// TwinCAT 3 PLC project MQTT_PLC_TEST
// ProgramVersion: 3.1.4024.0
// libraries:
//   Tc2_Standard, * (Beckhoff Automation GmbH)
//   Tc2_System, * (Beckhoff Automation GmbH)
//   Tc2_Utilities, * (Beckhoff Automation GmbH)
//   Tc3_IotBase, * (Beckhoff Automation GmbH)
//   Tc3_Module, * (Beckhoff Automation GmbH)
// project tree:
//   / GlobalTextList.TcGTLO, PlcTask.TcTTO
//   GVLs/ GVL_Visu.TcGVL, GVL_Mqtt.TcGVL
//   POUs/ MAIN.TcPOU
//   VISUs/ PannenkoekenDashboard.TcVIS
// real-time tasks:
//   TASK PlcTask: cycle T#10ms, priority 20, ADS port 350
// I/O:
//   DEVICE Device 1 (EtherCAT) (disabled), AmsNetId 199.4.42.250.2.1
//     Term 1 (EK1200) [EK1200-5000 EtherCAT Power supply (2A E-Bus)]
//       Term 2 (EL1008) [EL1008 8Ch. Dig. Input 24V, 3ms]
//       Term 3 (EL2008) [EL2008 8Ch. Dig. Output 24V, 0.5A]
//       Term 4 (EL3062) [EL3062 2Ch. Ana. Input 0-10V]
//       Term 5 (EL4002) [EL4002 2Ch. Ana. Output 0-10V, 12bit]
//       Term 6 (EK1110) [EK1110 EtherCAT extension]

CONFIGURATION MQTT_PLC_TEST
    RESOURCE PLC ON TwinCAT3
        TASK PlcTask(INTERVAL := T#10ms, PRIORITY := 20);
        PROGRAM MAIN WITH PlcTask : MAIN;
    END_RESOURCE
END_CONFIGURATION

// ---- GVLs/GVL_Visu.TcGVL
{attribute 'qualified_only'}
VAR_GLOBAL
    // Robot Arm
    sRobotState        : STRING(10);   // idle, moving, error
    nRobotColor        : DWORD;        // kleur voor rectangle/LED
    bRobotCmdSentPulse : BOOL;         // pulse indicator
    bRobotStateParseError : BOOL;      // parse fout indicator
END_VAR

// ---- GVLs/GVL_Mqtt.TcGVL
VAR_GLOBAL CONSTANT
    c_sMqttHost           : STRING(63) := '192.168.0.197';
    c_nMqttPort           : UINT := 1883;

    c_sTopicRobotCmd      : STRING(127) := 'pancake/robot/cmd';
    c_sTopicRobotState    : STRING(127) := 'pancake/robot/state';
    c_sTopicRobotError    : STRING(127) := 'pancake/robot/error';
    c_sTopicConveyorCmd   : STRING(127) := 'pancake/conveyor/cmd';
    c_sTopicConveyorState : STRING(127) := 'pancake/conveyor/state';
    c_sTopicConveyorError : STRING(127) := 'pancake/conveyor/error';
END_VAR

VAR_GLOBAL
    bMqttEnable                : BOOL := TRUE;
    bMqttConnected             : BOOL;
    bMqttError                 : BOOL;
    sMqttStatus                : STRING(127);

    sRobotState                : STRING(31) := 'unknown';
    bRobotStateUpdated         : BOOL;
    bRobotStateParseError      : BOOL;

    sConveyorCmdRx             : STRING(31);
    bConveyorCmdUpdated        : BOOL;
    sConveyorState             : STRING(31) := 'stopped';
    sConveyorStatePublished    : STRING(31);
    bConveyorStateSentPulse    : BOOL;
    sConveyorErrorText         : STRING(127);
    bConveyorErrorSentPulse    : BOOL;
    sConveyorItem              : STRING(31);
    bConveyorItemPresent       : BOOL;
    bConveyorItemUpdated       : BOOL;

    sRobotErrorRx              : STRING(127);
    bRobotErrorUpdated         : BOOL;

    sRobotCmdRequest           : STRING(31);
    bRobotCmdRequestPulse      : BOOL;
    sRobotCmdPending           : STRING(31);
    sRobotCmdSent              : STRING(31);
    bRobotCmdSentPulse         : BOOL;

    sCoordinatorState          : STRING(31);
    sLastRxTopic               : STRING(127);
    sLastRxPayload             : STRING(255);

    bCmdPick                   : BOOL;
    bCmdPlace                  : BOOL;
    bCmdHome                   : BOOL;
    bCmdStop                   : BOOL;
END_VAR

// ---- POUs/MAIN.TcPOU
PROGRAM MAIN
VAR
END_VAR

END_PROGRAM

// ---- GlobalTextList.TcGTLO
TEXTLIST GlobalTextList
  14 = 'Broker Host'
  78 = 'Broker Port'
  184 = 'Connected'
  631 = 'E-STOP'
  815 = 'E-STOPS'
  297 = 'Enable MQTT'
  818 = 'Error'
  717 = 'Mixer'
  369 = 'MQTT Broker'
  28 = 'MQTT Monitor'
  441 = 'Robot Arm'
  964 = 'Robot State'
  282 = 'S'
  632 = 'Status'
  865 = 'Transportband'
END_TEXTLIST

// ---- VISUs/PannenkoekenDashboard.TcVIS
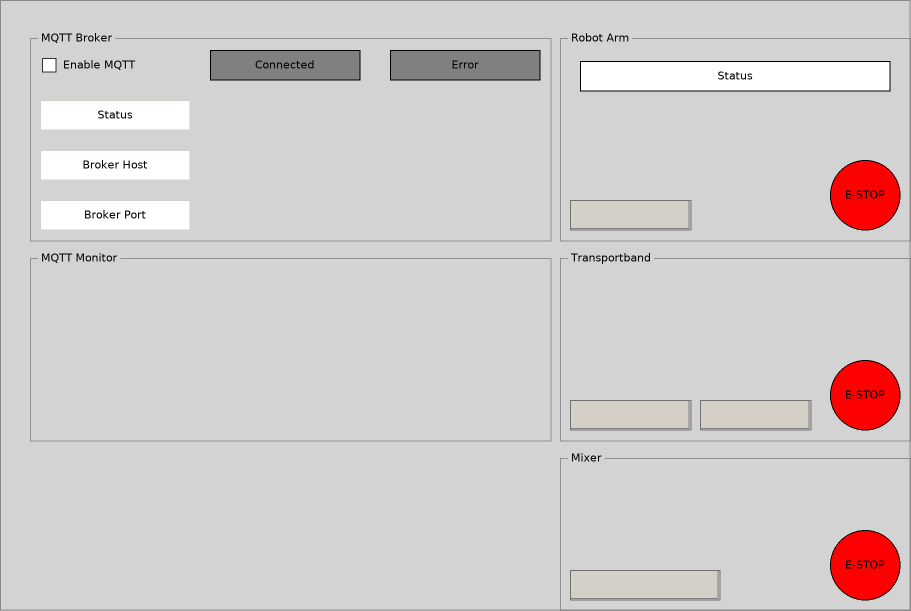
VISUALIZATION PannenkoekenDashboard  // 911x611
    GroupBox (30,30 521x211), "MQTT Broker"
        Checkbox (10,20 150x30), "Enable MQTT"
        Rectangle (360,20 150x30), "Error"
        Rectangle (180,20 150x30), "Connected"
        Textfield (10,70 150x30), "Status"
        Textfield (10,120 150x30), "Broker Host"
        Textfield (10,170 150x30), "Broker Port"
    GroupBox (30,250 521x191), "MQTT Monitor"
    GroupBox (560,30 351x211), "Robot Arm"
        Rectangle (20,31 310x30), "Status"
        Ellipse (270,130 70x70), "E-STOP"
        Button (10,170 121x30)
    GroupBox (560,250 351x191), "Transportband"
        Ellipse (270,110 70x70), "E-STOP"
        Button (10,150 121x30)
        Button (140,150 111x30)
    GroupBox (560,450 351x161), "Mixer"
        Ellipse (270,80 70x70), "E-STOP"
        Button (10,120 150x30)
END_VISUALIZATION
